{region 'Documentation'}
(*!
<summary>Checks equality with the expected SINT value.</summary>
*)
{endregion}
FUNCTION_BLOCK AssertEqual_SInt EXTENDS AssertionBase
VAR_INPUT
    IN : SINT; //! Actual value checked or observed by this Assertion.
    Expected : SINT; //! Reference value for comparison with IN.
END_VAR

SUPER^();

{region 'Documentation'}
(*!
<summary>Check equality with the expected SINT value.</summary>
*)
{endregion}
METHOD PROTECTED Assert
VAR
    Message : STRING(GVL_Constants.MessageLength);
    ExpectedText : STRING(GVL_Constants.AssertionValueLength);
    ActualText : STRING(GVL_Constants.AssertionValueLength);
END_VAR
IF NOT EvaluationActive THEN
    RETURN;
END_IF;

IF Result = E_Result.Error THEN
    RETURN;
END_IF;

IF Result = E_Result.Failed THEN
    RETURN;
END_IF;

IF IN <> Expected THEN
    ExpectedText := SINT_TO_STRING(Expected);
    ActualText := SINT_TO_STRING(IN);
    Message := CONCAT('Assertion failed: values are not equal. Expected = ',
        ExpectedText);
    Message := CONCAT(Message, ', Actual = ');
    Message := CONCAT(Message, ActualText);
    Message := CONCAT(Message, '.');
    Fail(Message := Message);
    RETURN;
END_IF;

Pass();
END_METHOD

END_FUNCTION_BLOCK

(* stored: Version 1.1.0.1
   POU AssertEqual_SInt: Id {0dae4e72-a5fa-4f3f-a5de-053cbbddd43c}, SpecialFunc None
   Folder Internal: Id {0880af0e-c030-4e17-948e-8c3877ccf26b}
   Method Assert: Id {4f79c20e-9a6d-42a1-b99a-62f090da909e} *)
